// TIA Portal V21 export
// export: Created 2026-11-21T13:26:58.8442366Z, ExportSetting WithDefaults, DisplayName Totally Integrated Automation Portal, DisplayVersion V21, DisplayName STEP 7 Professional, DisplayVersion V21, DisplayName STEP 7 Safety, DisplayVersion V21, DisplayName Tech WebApplication, DisplayVersion V21, DisplayName WinCC Basic/Comfort/Advanced, DisplayVersion V21, DisplayName WinCC Unified, DisplayVersion V21
FUNCTION_BLOCK "Valve"   // FB20, LAD
TITLE = Ventil / Valve / Vanne
{ S7_Optimized_Access := 'TRUE' }
VERSION : 0.1
// Ein Ventil mit Rückmeldung. / A valve with feedback. / Une vanne avec retour d'information.
// stored: AutoNumber true, IsIECCheckEnabled false, IsRetainMemResEnabled false, MemoryReserve 100, SetENOAutomatically false, UDAEnableTagReadback false
   VAR_INPUT
      open : Bool;   // Ventil öffnen / Open the valve / Ouvrir la vanne
      close : Bool;   // Close the valve
   END_VAR
   VAR_OUTPUT
      opened : Bool;   // Vanne ouverte
   END_VAR
   VAR
      moving : Bool;   // Ventil fährt / Valve is moving / La vanne se déplace
   END_VAR
BEGIN

REGION Network 1: Öffnen / Open / Ouvrir
   // Öffnen setzt das Fahren. / Opening starts the travel. / L'ouverture lance le déplacement.
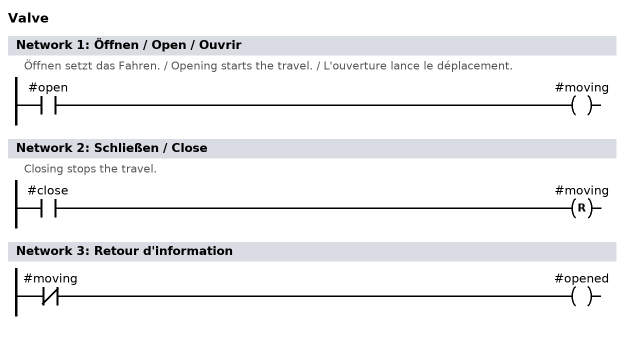
   RUNG wire#powerrail
      Contact( #open )
      Coil( #moving )
   END_RUNG
   // the same network as SCL:
   #moving := #open;
END_REGION

REGION Network 2: Schließen / Close
   // Closing stops the travel.
   RUNG wire#powerrail
      Contact( #close )
      R_Coil( #moving )
   END_RUNG
   // the same network as SCL:
   IF #close THEN #moving := FALSE; END_IF;
END_REGION

REGION Network 3: Retour d'information
   RUNG wire#powerrail
      I_Contact( #moving )
      Coil( #opened )
   END_RUNG
   // the same network as SCL:
   #opened := NOT #moving;
END_REGION
END_FUNCTION_BLOCK
